Fanuc KAREL source: kt00294.KL

-- PROVISIONAL review KL for V770-1; original PC SHA256 713b76724aa8cb3113ee6a2b200c2bc2189fb1da18e7a8ccd343a4f6caad909e
-- Incomplete behavior may be omitted. Consult companion uncertainty JSON. Do not deploy.
PROGRAM KT00294
%NOLOCKGROUP
VAR
  I1 : INTEGER
  R2 : REAL
  OUT : BOOLEAN
BEGIN
  -- UNRESOLVED_PC offsets 5-16; opcodes 2E,23
  -- UNRESOLVED_PC offsets 21-32; opcodes 2E,23
  -- UNRESOLVED_PC offsets 37-58; opcodes 21,21,29,64,6E,23
  -- UNRESOLVED_PC offsets 63-67; opcodes 7F
END KT00294
